(* IEC 61131-3 sources: IRIS-Project/LASAL CONTROL SOFTWARE/LasalProject_2025_09_12/Class/SafetyManager (part 6) *)

    sUdpVars.CalculatedRequestTimeout := Temp;
    bGetRequestTimeout := TRUE;
  else
    // activate the default settings (min settings)
    sUdpVars.CalculatedRequestTimeout := UDP_MIN_REQUEST_TIMEOUT;
  end_if;

  // use default value for request time
  sUdpVars.CalculatedRequestTime    := UDP_MIN_REQUEST_TIME;

  //check for advanced request time from user
  if sUdpVars.udAdvancedRequestCycle >= UDP_MIN_REQUEST_TIME
  & sUdpVars.udAdvancedRequestCycle <= (sUdpVars.CalculatedRequestTimeout/2)  then
    sUdpVars.CalculatedRequestTime := sUdpVars.udAdvancedRequestCycle;
  else
    //only log error if we got calculated request timeout and value is not zero
    if bGetRequestTimeout = TRUE & sUdpVars.udAdvancedResponseTimeout <> 0 & bd_SingleLog.SetUdpRequestCycleFailed = FALSE then
      LogValue("@04D6 (SafetyManager::SetUdpSchedulerGrid) [SL] The value of 0x{0} for the UDP Request Cycle is not valid! The maximum value is 0x{1}", Value:=sUdpVars.udAdvancedRequestCycle, (sUdpVars.CalculatedRequestTimeout/2));
      bd_SingleLog.SetUdpRequestCycleFailed := TRUE;
    end_if;
  end_if;

  // always use the min settings for the responses
  sUdpVars.CalculatedResponseTime    := UDP_MIN_RESPONSE_TIME;
  sUdpVars.CalculatedResponseTimeout := UDP_MIN_RESPONSE_TIMEOUT;

  //check for advanced response timeout from user
  if sUdpVars.udAdvancedResponseTimeout >= UDP_MIN_RESPONSE_TIMEOUT then
    sUdpVars.CalculatedResponseTimeout := sUdpVars.udAdvancedResponseTimeout;
  else
    // only log error if value is not zero
    if sUdpVars.udAdvancedResponseTimeout <> 0 & bd_SingleLog.SetUdpResponseTimeoutFailed = FALSE then
      LogValue("@04D7 (SafetyManager::SetUdpSchedulerGrid) [SL] The value of 0x{0} for the UDP Response Timeout is not valid! The minimum value is 0x{1}", Value:=sUdpVars.udAdvancedResponseTimeout, UDP_MIN_RESPONSE_TIMEOUT);
      bd_SingleLog.SetUdpResponseTimeoutFailed := TRUE;
    end_if;
  end_if;

END_FUNCTION

FUNCTION SafetyManager::UdpResponseScheduler
  VAR
    pActResponseEntry : ^t_UdpConnection;
    pActRetryEntry    : ^t_UdpConnection;
    tmpretcode        : DINT;
    i                 : UDINT;
  END_VAR

  //point to actual request-entry
  pActResponseEntry := #sUdpVars.paConnectionsToConsumers^[sUdpVars.ResponseScheduler.ActRequestedIndex];

  //send a request every TRequestTime x Cycnt Cycle
  if ((sUdpVars.ResponseScheduler.CyCnt MOD sUdpVars.CalculatedResponseTime) = 0) then

    // search through the list if something has to be sent (check also for changes in the data)
    for i := 0 to sUdpVars.ConsumerConnectionNo-1 do

      //only send a request if not waiting for a response and the IP is valid (on cleaning out the connections some may be set to 0)
      if (pActResponseEntry^.WaitForResponse = FALSE) & (pActResponseEntry^.IP <> 0) & (pActResponseEntry^.SendResponse = TRUE) then

        //send request to mover of actual entry
        tmpretcode := SendUdpResponse(pActResponseEntry);
        if tmpretcode >= 0 then

          //if sending was successful we are waiting for a response
          pActResponseEntry^.WaitForResponse := TRUE;
          pActResponseEntry^.SendResponse    := FALSE;
          pActResponseEntry^.TLastRequest      := ops.tAbsolute;
          pActResponseEntry^.RequestRetries    := 0;

        else
          //unable to send request
          if bd_SingleLog.SendUdpRspFailed = FALSE then
            bd_SingleLog.SendUdpRspFailed := TRUE;
            LogError("@04A0 (SafetyManager::UdpResponseScheduler) [SL] Failed to send udp response");
          end_if;
        end_if;

      end_if;

      //increase actual index
      if sUdpVars.ResponseScheduler.ActRequestedIndex < (sUdpVars.ConsumerConnectionNo-1) then
        sUdpVars.ResponseScheduler.ActRequestedIndex += 1;
      else
        //when reaching last entry -> reset index
        sUdpVars.ResponseScheduler.ActRequestedIndex := 0;
      end_if;

      pActResponseEntry := #sUdpVars.paConnectionsToConsumers^[sUdpVars.ResponseScheduler.ActRequestedIndex];
    end_for;

  // between the normal requests we do the retries
  elsif ((sUdpVars.ResponseScheduler.CyCnt MOD UDP_RETRY_TIME) = 0) then

    pActRetryEntry := #sUdpVars.paConnectionsToConsumers^[0];

    // check if we have to send a retry
    for i := 0 to sUdpVars.ConsumerConnectionNo-1 do

      // look if we actual wait for a response to send retries and check if we didn't receive data in time
      if (pActRetryEntry^.WaitForResponse = TRUE) & ((ops.tAbsolute - pActRetryEntry^.TLastRequest) > sUdpVars.CalculatedResponseTimeout) then

        if pActRetryEntry^.RequestRetries >= UDP_MAX_RETRIES then

          pActRetryEntry^.MaxRetryCnt          += 1;
          pActRetryEntry^.WaitForResponse      := FALSE;
          //don't reset flag here, because it's possible we receive an old sequence counter with next package, which leads to an error at FSoE communication
          //pActRetryEntry^.bSequenceCntReceived := FALSE; //reset flag to allow sequence counter for new udp communication

        // only if the IP is valid
        elsif (pActRetryEntry^.IP <> 0) then

          //send retry to actual cpu
          tmpretcode := SendUdpResponse(pActRetryEntry);
          if tmpretcode >= 0 then
            pActRetryEntry^.TLastRequest   := ops.tAbsolute;
            pActRetryEntry^.RequestRetries += 1;
            exit;
          else
            //unable to send retry
            if bd_SingleLog.SendUdpRspRetryFailed = FALSE then
              bd_SingleLog.SendUdpRspRetryFailed := TRUE;
              LogError("@049D (SafetyManager::UdpResponseScheduler) [SL] Failed to send udp retry");
            end_if;
          end_if;
        end_if;

      end_if;

      pActRetryEntry += sizeof(t_UdpConnection);

    end_for;

  end_if;

  sUdpVars.ResponseScheduler.CyCnt += 1;

END_FUNCTION

FUNCTION SafetyManager::SendUdpResponse
  VAR_INPUT
    pConnection 	: ^t_UdpConnection;
  END_VAR
  VAR_OUTPUT
    retcode 	: DINT;
  END_VAR
  VAR
    udActSendLength : UDINT;
  END_VAR

  sUdpVars.pTempSendBufferCy^.Header.Command   := t_UdpCommand::UdpCmd_DataRsp;
  //The current header version is set here so that the other side knows which version is supported.
  sUdpVars.pTempSendBufferCy^.Header.State     := t_UdpPacketHeaderV2.State.IsFromProducer + UDP_HEADER_ACTVERSION;
  sUdpVars.pTempSendBufferCy^.Header.IFCRC     := pConnection^.IFCRC;
  sUdpVars.pTempSendBufferCy^.Header.SafetyNbr := pConnection^.SafetyNbr;

  UdpSendData.SectionStart();

  //check for new header version with extended sequence number (4Byte)
  if pConnection^.ActSendData.usHeaderVersion >= UDP_HEADER_VERSION_V2 then

    sUdpVars.pTempSendBufferCy^.Header.SequenceNumber := pConnection^.ActSendData.udSequenceNumber;

    udActSendLength := sizeof(t_UdpPacketHeaderV2);

    if pConnection^.ActSendData.PdoLength then
      sUdpVars.pTempSendBufferCy^.Header.PdoDataLength  := pConnection^.ActSendData.PdoLength;
      _memcpy(ptr1:=#sUdpVars.pTempSendBufferCy^.Data, ptr2:=#pConnection^.ActSendData.PdoData, cntr:=pConnection^.ActSendData.PdoLength);
      udActSendLength += pConnection^.ActSendData.PdoLength;
    else
      sUdpVars.pTempSendBufferCy^.Header.PdoDataLength  := 0;
    end_if;

    if pConnection^.ActSendData.SdoLength then
      sUdpVars.pTempSendBufferCy^.Header.SdoDataLength  := pConnection^.ActSendData.SdoLength;
      _memcpy(ptr1:=#sUdpVars.pTempSendBufferCy^.Data + pConnection^.ActSendData.PdoLength, ptr2:=#pConnection^.ActSendData.SdoData, cntr:=pConnection^.ActSendData.SdoLength);
      udActSendLength += pConnection^.ActSendData.SdoLength;
    else
      sUdpVars.pTempSendBufferCy^.Header.SdoDataLength  := 0;
    end_if;
  else
    //use old headerversion with 1byte Sequence Counter
    sUdpVars.pTempSendBufferCy^$t_UdpPacketV1.Header.SequenceNumber := pConnection^.ActSendData.usSequenceNumber;

    udActSendLength := sizeof(t_UdpPacketHeaderV1);

    if pConnection^.ActSendData.PdoLength then
      sUdpVars.pTempSendBufferCy^$t_UdpPacketV1.Header.PdoDataLength  := pConnection^.ActSendData.PdoLength;
      _memcpy(ptr1:=#sUdpVars.pTempSendBufferCy^$t_UdpPacketV1.Data, ptr2:=#pConnection^.ActSendData.PdoData, cntr:=pConnection^.ActSendData.PdoLength);
      udActSendLength += pConnection^.ActSendData.PdoLength;
    else
      sUdpVars.pTempSendBufferCy^$t_UdpPacketV1.Header.PdoDataLength  := 0;
    end_if;

    if pConnection^.ActSendData.SdoLength then
      sUdpVars.pTempSendBufferCy^$t_UdpPacketV1.Header.SdoDataLength  := pConnection^.ActSendData.SdoLength;
      _memcpy(ptr1:=#sUdpVars.pTempSendBufferCy^$t_UdpPacketV1.Data + pConnection^.ActSendData.PdoLength, ptr2:=#pConnection^.ActSendData.SdoData, cntr:=pConnection^.ActSendData.SdoLength);
      udActSendLength += pConnection^.ActSendData.SdoLength;
    else
      sUdpVars.pTempSendBufferCy^$t_UdpPacketV1.Header.SdoDataLength  := 0;
    end_if;

  end_if;

  UdpSendData.SectionStop();

  retcode := SendUDPData(sUdpVars.pTempSendBufferCy, udActSendLength, pConnection^.IP);

  sUdpVars.SendCnt += 1;

  if retcode < 0 then
    // error at sending
    sUdpVars.LastSendError := retcode;
    sUdpVars.SendErrorCnt += 1;
  else
    // only valid one-time
    pConnection^.ActSendData.SdoLength    := 0;

    pConnection^.SentPackages += 1;
  end_if;

END_FUNCTION

FUNCTION SafetyManager::UdpTask

  while TRUE do

        // if there is no error and we got UDP stuff going on => do it
    if (sUdpVars.ProducerConnectionNo | ((sUdpVars.UdpInit AND 2#11) = (t_UdpInit.FSoEAvailable OR t_UdpInit.ProvidesIF))) then
      if sUdpVars.UdpInit.CallBackInstalled = FALSE then

        //add callback info for receiving udp packages
        AddCallBackInfo(this, #ReceiveUDPData());

        sUdpVars.UdpInit.CallBackInstalled := TRUE;
      end_if;

      SafetyUDP::CyWork(0);

      // no SDOs or scheduling when we reinitialize
      if CommInitialized & (InitSSW > _ClearRoutingInfos) then
        // check initialisation of the connections
        if sUdpVars.ConnectionsInitialized = FALSE then
          ShareUdpConnectionInfos();
        end_if;

        // only if we're a consumer and have producers to contact
        if sUdpVars.ProducerConnectionNo then

          // work the connections (send requests)
          UdpRequestScheduler();

          // forward the SDOs from the producer (responses)
          ForwardReceivedUdpSDOs(paConnections:=sUdpVars.paConnectionsToProducers, ConnectionNo:=sUdpVars.ProducerConnectionNo);
        end_if;

        // if there are consumers, we may distribute new SDO data
        if sUdpVars.ConsumerConnectionNo then

          // work the connections (send responses)
          UdpResponseScheduler();

          // forward the SDOs from the consumers (requests)
          ForwardReceivedUdpSDOs(paConnections:=sUdpVars.paConnectionsToConsumers, ConnectionNo:=sUdpVars.ConsumerConnectionNo);
        end_if;
      end_if;
    end_if;

    To_MultiTask.TASKDELAY(timeout0:=1);
  end_while;

END_FUNCTION

FUNCTION SafetyManager::TimeSyncModuleAvailable
  VAR_INPUT
    pTimeSyncElement 	: ^t_TimeSyncElement;
  END_VAR
  VAR_OUTPUT
    Available 	: BOOL;
  END_VAR

  if pTimeSyncElement^.InfoBits.IsMissingOptional | (pTimeSyncElement^.pSafety & (pTimeSyncElement^.pSafety^.SafetyNbr = 0)) then
    Available := FALSE;
  else
    Available := TRUE;
  end_if;

END_FUNCTION

FUNCTION SafetyManager::ReinitEverything
  VAR
    MyPara 	  : CmdStruct;
    MyResult 	: results;
  END_VAR

  // new safety project detected (different crc) => reinit the system (similar to disconnect)
  MyPara.uiCmd := CMD_SM_DISCONNECT;
  MyPara.aPara[0] := 0; // set length of further parameters to 0
  TellAllInterfaceManagingModules(#MyPara, #MyResult);  // tell all interface domains to reestablish connection (they need the safety number from the configuration)
  TellAllSafetyModules(#MyPara, #MyResult);             // tell all of our local safety modules that there's a new config => reinitialize

  ClassState := 0;

  // reset module sync no (no more modules synchron)
  ModuleSyncNo := 0;

  // restart initialisation (maybe we had no clue about interfaceframes when initialising the first time)
  InitSSW := _ClearRoutingInfos;

END_FUNCTION

FUNCTION SafetyManager::CheckCustomConnectionValid
  VAR_INPUT
    pConnection 	: ^t_FSoEConnectionDetails;
    pIFFSoEInfo 	: ^t_FSoEConnInfo;
  END_VAR
  VAR_OUTPUT
    bIsCustomConnValid 	: BOOL;
  END_VAR

  // This method checks if the passed connection and FSoE Interface are a Valid custom connection
  // This check replaces the slave address check for normal FSoE Interface frames. (s. FinalizePDOMapping)
  // (The slave addresses may not valid for custom connections at this point)

  bIsCustomConnValid := FALSE;

  if pConnection = NIL | pIFFSoEInfo = NIL | pIFFSoEInfo^.pManaging = NIL then
    return;
  end_if;

  if pConnection^.Flags.IsMaster then

    // Check for custom ip address in compressed path
    // Check for HWT_ESCAPE_SAFETY_CUSTOM in uncompressed path
    // pConnection^.pSlavePathComp: 1 Byte Type, 4 Byte IF CRC, 4 Byte Custom IP Addr,
    // example : 03 59 8C AE 3D 00 00 00 02 FF FF FF
    // pIFFSoEInfo^.pManaging^.pModulePath: 2 Byte Length, 1 Byte Domain No, 1 Byte Escape Sequence, 1 Byte Custom IP Addr
    // example : 03 00 00 8A 02
    if pConnection^.pSlavePathComp & pConnection^.SlavePathCompLen > 8 &                    // Pointer + length (Custom IP = Byte 9)
       (pConnection^.pSlavePathComp^ = 3) &                                                 // Type Code
       pIFFSoEInfo^.pManaging^.pModulePath & (pIFFSoEInfo^.pManaging^.pModulePath^ >= 3) &  // Pointer + length
       ((pConnection^.pSlavePathComp+5)^$UDINT AND 16#00FFFFFF) = 0 &                       // Custom IP
       (pIFFSoEInfo^.pManaging^.pModulePath+3)^ = HWT_ESCAPE_SAFETY_CUSTOM  then            // Escape Sequence
      // Compare Custom IDs
      if (pConnection^.pSlavePathComp + 8)^ = (pIFFSoEInfo^.pManaging^.pModulePath+4)^ then
        bIsCustomConnValid := TRUE;
      end_if;

    end_if;

  else

    // Check IFCRC in compressed path
    // Check for HWT_ESCAPE_SAFETY_CUSTOM in uncompressed path
    // pConnection^.pSlavePathComp: 1 Byte Type, 4 Byte IF CRC
    // example : 03 59 8C AE 3D FF FF FF
    // pIFFSoEInfo^.pManaging^.pModulePath: 2 Byte Length, 1 Byte Domain No, 1 Byte Escape Sequence, 1 Byte Custom IP Addr
    // example : 03 00 00 8A 02
    if pConnection^.pSlavePathComp & pConnection^.SlavePathCompLen > 5 &                    // Pointer + length (IFCRC = Byte 1, 4Byte CRC Data )
       (pConnection^.pSlavePathComp^ = 3) &                                                 // Type Code
       pIFFSoEInfo^.pManaging^.pModulePath & (pIFFSoEInfo^.pManaging^.pModulePath^ >= 3) &  // Pointer + length
       (pIFFSoEInfo^.pManaging^.pModulePath+3)^ = HWT_ESCAPE_SAFETY_CUSTOM then             // Escape Sequence

      // Compare IFCRC (Cannot compare Custom IDs because (pConnection^.pSlavePathComp + 8)^ may not be valid yet at this time
      if (pConnection^.pSlavePathComp+1)^$UDINT = pIFFSoEInfo^.FromOtherSide.InterfaceCRC then
        bIsCustomConnValid := TRUE;
      end_if;

    end_if;

  end_if;

END_FUNCTION

FUNCTION SafetyManager::ShareSingleConnectionInfos
	VAR_INPUT
		pMasterConnection 	: ^t_FSoEConnectionDetails;
		pModuleConfig 	: ^t_ModuleListElem;
	END_VAR
  VAR
  	pMasterModuleCfg  : ^t_ModuleListElem;
  	pSlaveModuleCfg   : ^t_ModuleListElem;
    pActModuleCfg     : ^t_ModuleListElem;
    pHelpSafety       : ^t_SafetyComponent;
    pMasterSafety     : ^t_SafetyComponent;
    pSlaveSafety      : ^t_SafetyComponent;
    MyPara 	          : CmdStruct;
    MyResult	        : results;
    pPDOReadData      : pVoid;
    i                 : UDINT;
    IsInList          : BOOL;
  END_VAR

//*****************************************************************************
//** TELL THE MODULES WHAT DATA TO COPY IN REALTIME                          **
//*****************************************************************************

  // get the master and slave module configuration of this connection

  // master module configuration is always the first one in the list
  pMasterModuleCfg  := pModuleConfig;

  // search for the slave config via the path stored in the connection
  pSlaveModuleCfg   := NIL;
  pActModuleCfg     := pModuleConfig;
  while pActModuleCfg do
    if (pActModuleCfg^.ModuleInfo.pPath^ = pMasterConnection^.pSlavePath^) &
       (To_StdLib.MemCmp(pActModuleCfg^.ModuleInfo.pPath+1, pMasterConnection^.pSlavePath+1, pMasterConnection^.pSlavePath^+1) = 0) then

      pSlaveModuleCfg := pActModuleCfg;
      exit;
    end_if;

    pActModuleCfg := pActModuleCfg^.pNext;
  end_while;

  if pSlaveModuleCfg = NIL then
    return;
  end_if;

  // get the object this pointers via the hardware paths
  pMasterSafety := NIL;
  pSlaveSafety  := NIL;

  pHelpSafety := pFirstSafetyComponent;
  while pHelpSafety do
    if pHelpSafety^.PathLen &
       (pMasterModuleCfg^.ModuleInfo.pPath^ = pHelpSafety^.pPath^) &
       (To_StdLib.MemCmp(pHelpSafety^.pPath + 1, pMasterModuleCfg^.ModuleInfo.pPath + 2 + pMasterModuleCfg^.ModuleInfo.pPath^ - pHelpSafety^.pPath^, pHelpSafety^.pPath^) = 0) then
      pMasterSafety := pHelpSafety;
      exit;
    else
      pHelpSafety := pHelpSafety^.pNext;
    end_if;
  end_while;

  pHelpSafety := pFirstSafetyComponent;
  while pHelpSafety do
    if pHelpSafety^.PathLen &
       (pSlaveModuleCfg^.ModuleInfo.pPath^ = pHelpSafety^.pPath^) &
       (To_StdLib.MemCmp(pHelpSafety^.pPath + 1, pSlaveModuleCfg^.ModuleInfo.pPath + 2 + pSlaveModuleCfg^.ModuleInfo.pPath^ - pHelpSafety^.pPath^, pHelpSafety^.pPath^) = 0) then
      pSlaveSafety := pHelpSafety;
      exit;
    else
      pHelpSafety := pHelpSafety^.pNext;
    end_if;
  end_while;

  if pMasterSafety & pSlaveSafety then

    // we start with the safe outputs: get the data pointer from the master and give it to the slave
    MyPara.uiCmd    := CMD_SM_ADD_OUTPUT_PDO;
    MyResult.uiLng  := 0;
    pMasterSafety^.pThis^.NewInst(#MyPara, #MyResult);

    if MyResult.uiLng <> 4 then
      LogError("@048F (SafetyManager::ShareSingleConnectionInfos) Invalid return value when asking the master safety module for it's pointer to the PDO read data!");
      return;
    end_if;

    pPDOReadData := MyResult.aData[0]$pVoid;

  #ifdef SAFETY_DEBUG_LOGGING_ACTIVATED
  #pragma message("RamAnd 20.11.2014 16:41 \ testweise mapping loggen")
    LogValue("@DBG (SafetyManager::ShareSingleConnectionInfos) ConnectionID: {0}, SlaveAddress: {1}", Value:=pMasterConnection^.ConnectionID, Value2:=pMasterConnection^.SlaveAddress);
    LogValue("@DBG (SafetyManager::ShareSingleConnectionInfos) MasterSafetyNbr: {0}, SlaveSafetyNbr: {1}", Value:=pMasterSafety^.SafetyNbr, Value2:=pSlaveSafety^.SafetyNbr);
    LogValue("@DBG (SafetyManager::ShareSingleConnectionInfos) MasterReadOffset: {0}, MasterReadSize: {1}, SlaveWriteOffset: {2}", Value:=pMasterConnection^.MasterReadOffset, Value2:=pMasterConnection^.MasterReadSize, Value3 := pMasterConnection^.SlaveWriteOffset);
  #endif

    // check if it's in the list
    IsInList := FALSE;
    if FSoEInputPDONo then
      for i := 0 to (FSoEInputPDONo-1) do
        if ((aFSoEInputPDOs[i].pSafety = pSlaveSafety)  & (aFSoEInputPDOs[i].pMem = pPDOReadData$DINT + pMasterConnection^.MasterReadOffset)) then
          aFSoEInputPDOs[FSoEInputPDONo].pSafety    := pMasterSafety;
          aFSoEInputPDOs[FSoEInputPDONo].pMem       := MyPara.aPara[0];
          IsInList := TRUE;
        end_if;
      end_for;
    end_if;

    if IsInList = FALSE then
      MyPara.uiCmd    := CMD_SM_ADD_INPUT_PDO;
      MyPara.aPara[0] := pPDOReadData$DINT + pMasterConnection^.MasterReadOffset;
      MyPara.aPara[2] := pMasterConnection^.OwnerSafetyNbr$DINT;
      MyPara.aPara[3] := pMasterConnection^.MasterReadSize;
      MyPara.aPara[4] := pMasterSafety^.InfoBits.IsOptional;
      MyPara.aPara[7] := pMasterConnection^.SlaveWriteOffset;
      MyPara.aPara[8] := SM_IF_VALIDITY_MARK$DINT;
      MyPara.aPara[9] := pMasterConnection^.Flags.IsInterfaceConnection;
      pSlaveSafety^.pThis^.NewInst(#MyPara, #MyResult);

      if FSoEInputPDONo < MAX_FSOE_CONNECTIONS then
        aFSoEInputPDOs[FSoEInputPDONo].pSafety    := pSlaveSafety;
        aFSoEInputPDOs[FSoEInputPDONo].pMem       := MyPara.aPara[0];
        FSoEInputPDONo += 1;
      else
        LogValue("@0490 (SafetyManager::ShareSingleConnectionInfos) Maximum limit of allowed FSoE input Frames exceeded (0x{0})", Value:=MAX_FSOE_CONNECTIONS);
      end_if;
    end_if;

    // safe inputs: get the data pointer from the slave and give it to the master
    MyPara.uiCmd    := CMD_SM_ADD_OUTPUT_PDO;
    MyResult.uiLng  := 0;
    pSlaveSafety^.pThis^.NewInst(#MyPara, #MyResult);

    if MyResult.uiLng <> 4 then
      LogError("@0491 (SafetyManager::ShareSingleConnectionInfos) Invalid return value when asking the slave safety module for it's pointer to the PDO read data!");
      return;
    end_if;

    pPDOReadData := MyResult.aData[0]$pVoid;

  #ifdef SAFETY_DEBUG_LOGGING_ACTIVATED
  #pragma message("RamAnd 20.11.2014 16:41 \ testweise mapping loggen")
    LogValue("@DBG (SafetyManager::ShareSingleConnectionInfos) SlaveReadOffset: {0}, SlaveReadSize: {1}, MasterWriteOffset: {2}", Value:=pMasterConnection^.SlaveReadOffset, Value2:=pMasterConnection^.MasterWriteSize, Value3 := pMasterConnection^.MasterWriteOffset);
  #endif

    // check if it's in the list
    IsInList := FALSE;
    if FSoEInputPDONo then
      for i := 0 to (FSoEInputPDONo-1) do
        if ((aFSoEInputPDOs[i].pSafety = pMasterSafety)  & (aFSoEInputPDOs[i].pMem = pPDOReadData$DINT + pMasterConnection^.SlaveReadOffset)) then
          aFSoEInputPDOs[FSoEInputPDONo].pSafety    := pMasterSafety;
          aFSoEInputPDOs[FSoEInputPDONo].pMem       := MyPara.aPara[0];
          IsInList := TRUE;
        end_if;
      end_for;
    end_if;

    if IsInList = FALSE then

      MyPara.uiCmd    := CMD_SM_ADD_INPUT_PDO;
      MyPara.aPara[0] := pPDOReadData$DINT + pMasterConnection^.SlaveReadOffset;
      MyPara.aPara[2] := pSlaveSafety^.SafetyNbr$DINT;
      MyPara.aPara[3] := pMasterConnection^.MasterWriteSize;
      MyPara.aPara[4] := pSlaveSafety^.InfoBits.IsOptional;
      MyPara.aPara[7] := pMasterConnection^.MasterWriteOffset;
      MyPara.aPara[8] := 0;
      MyPara.aPara[9] := 0;
      pMasterSafety^.pThis^.NewInst(#MyPara, #MyResult);

      if FSoEInputPDONo < MAX_FSOE_CONNECTIONS then
        aFSoEInputPDOs[FSoEInputPDONo].pSafety    := pMasterSafety;
        aFSoEInputPDOs[FSoEInputPDONo].pMem       := MyPara.aPara[0];
        FSoEInputPDONo += 1;
      else
        LogValue("@0490 (SafetyManager::ShareSingleConnectionInfos) Maximum limit of allowed FSoE input Frames exceeded (0x{0})", Value:=MAX_FSOE_CONNECTIONS);
      end_if;
    end_if;

    // remember that we already dealt with this connection
    pMasterConnection^.InternalConnectionState := FCS_CONNECTION;

  end_if;

END_FUNCTION
